// SIMATIC S7-200 project (STEP 7-Micro/WIN), CPU 224 CN REL 02.01

SYMBOL_TABLE USUARIO1
SM2              I0.0     // Sensor magnetico extendido del cilindro retenedor
SM1              I0.1     // Sensor magnetico retraido del cilindor retenedor
SM4              I0.2     // Sensor magnetico extendido del cilindro de empuje
SM3              I0.3     // Sensor magnetico retraido del cilindor de empuje
SF               I0.4     // Sensor Fotoelectrico Final
SP               I0.5     // Sensor Fotoelectrico Superior
SP1              I0.6     // Sensor Fotoelectrico Inferior
SII              I0.7     // Sensor Inductivo
SB_1             I1.2     // Pulsador de marcha
SB_2             I1.3     // Pulsador de paro
QS               I1.4     // Zeta de Emergencia
SA               I1.5     // Selector de modo
KV1              Q0.0     // Cilindro neumatico Retenedor
KV2              Q0.1     // Cilindro neumatico de empuje
HL1              Q0.7     // Señalizacion amarillo
HL2              Q1.0     // Señalizacion verde
HL3              Q1.1     // Señalizacion roja
E0               M0.0     // Estado 0
E1               M0.1     // Estado 1
E2               M0.2     // Estado 2
E3               M0.3     // Estado 3
E4               M0.4     // Estado 4
E5               M0.5     // Estado 5
EM               M0.6     // Estado de emergencia
EP               M0.7     // Estado de parada
CONT1            VW270
END_SYMBOL_TABLE

ORGANIZATION_BLOCK PRINCIPAL:OB1
TITLE=COMENTARIOS DEL PROGRAMA
BEGIN
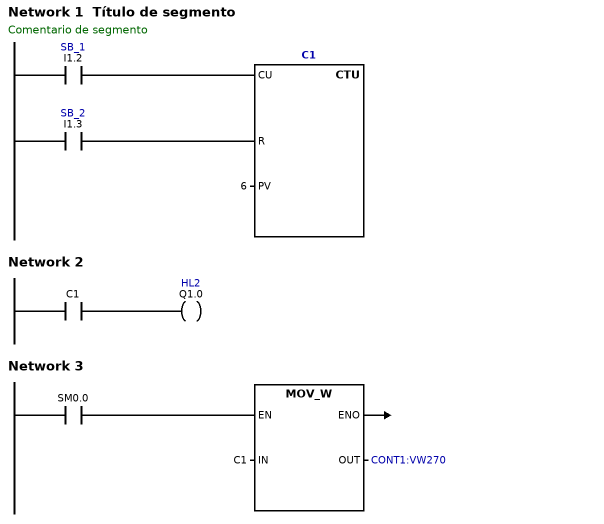
Network 1 // Título de segmento
// Comentario de segmento
LD     SB_1:I1.2
LD     SB_2:I1.3
CTU    C1, 6
Network 2
LD     C1
=      HL2:Q1.0
Network 3
LD     SM0.0
MOVW   C1, CONT1:VW270
END_ORGANIZATION_BLOCK
